(* IEC 61131-3 sources: plcassist-cli/packages/volt-lsp-iec/test-corpus/lenze-mid/Device/Plc Logic/Application/Library Manager/L_ILMP_LicenseManager, 13 files *)

(* ---- GETBOOLEANPROPERTY.fun ---- *)
FUNCTION GETBOOLEANPROPERTY : BOOL
VAR_INPUT
	STKEY : WSTRING;
END_VAR
END_FUNCTION

(* ---- GETCOMPANY.fun ---- *)
FUNCTION GETCOMPANY : WSTRING
END_FUNCTION

(* ---- GETNUMBERPROPERTY.fun ---- *)
FUNCTION GETNUMBERPROPERTY : DINT
VAR_INPUT
	STKEY : WSTRING;
END_VAR
END_FUNCTION

(* ---- GETTEXTPROPERTY.fun ---- *)
FUNCTION GETTEXTPROPERTY : WSTRING
VAR_INPUT
	STKEY : WSTRING;
END_VAR
END_FUNCTION

(* ---- GETTEXTPROPERTY2.fun ---- *)
FUNCTION GETTEXTPROPERTY2 : POINTER TO WSTRING
VAR_INPUT
	STKEY : WSTRING;
END_VAR
END_FUNCTION

(* ---- GETTITLE.fun ---- *)
FUNCTION GETTITLE : WSTRING
END_FUNCTION

(* ---- GETVERSION.fun ---- *)
FUNCTION GETVERSION : VERSION
END_FUNCTION

(* ---- GETVERSIONPROPERTY.fun ---- *)
FUNCTION GETVERSIONPROPERTY : VERSION
VAR_INPUT
	STKEY : WSTRING;
END_VAR
END_FUNCTION

(* ---- L_ILMP_LICENSECONFIGUPDATEFROMPLC.fun ---- *)
FUNCTION L_ILMP_LICENSECONFIGUPDATEFROMPLC : BOOL
END_FUNCTION

(* ---- L_ILMP_LICENSECONFIGUREMODE.fun ---- *)
FUNCTION L_ILMP_LICENSECONFIGUREMODE : DWORD
VAR_INPUT
	XUPDATE : BOOL;
	DWNEWCONFIGMODE : DWORD;
END_VAR
END_FUNCTION

(* ---- GLOBALTEXTLIST.fb ---- *)
FUNCTION_BLOCK GLOBALTEXTLIST
VAR
	M_TEXTLISTFILE : STRING(255);
	_STNAMESPACE : STRING;
END_VAR
END_FUNCTION_BLOCK

(* ---- L_ILMP_MANAGELICENSECONFIGURATION.fb ---- *)
FUNCTION_BLOCK L_ILMP_MANAGELICENSECONFIGURATION
VAR
	DWCONFIG : DWORD;
	APPLICATIONCREDITINFO : L_IMHP_LM_ApplicationCreditInfo;
	APPCREDITCONFIG : L_IMHP_LM_ApplicationCreditConfiguration;
END_VAR
END_FUNCTION_BLOCK

METHOD INITIALIZE : UDINT
VAR_INPUT
	WMODULETYPE : UINT;
	DWINSTANCE : UDINT;
	PCONNECTOR : POINTER TO IoConfigConnector;
END_VAR
END_METHOD

(* ---- L_ILMP_SETAPPCREDITCONFIGURATION.fb ---- *)
FUNCTION_BLOCK L_ILMP_SETAPPCREDITCONFIGURATION
VAR_INPUT
	XEXECUTE : BOOL;
	SCAPPCREDITCONFIG : L_ILMP_AppCreditConfiguration;
END_VAR
VAR_OUTPUT
	XBUSY : BOOL;
	XDONE : BOOL;
	XERROR : BOOL;
	EERRORID : L_ILMP_Error;
END_VAR
VAR
	XEXECUTEOLD : BOOL;
	DWCONFIG : DWORD;
	XBUSY_INT : BOOL;
	XDONE_INT : BOOL;
	APPLICATIONCREDITINFO : L_IMHP_LM_ApplicationCreditInfo;
	APPCREDITCONFIG : L_IMHP_LM_ApplicationCreditConfiguration;
END_VAR
END_FUNCTION_BLOCK

METHOD ABORT : UDINT
END_METHOD

METHOD EXECUTE : UDINT
END_METHOD
